TYPE "ST_StepRecord"
VERSION : 0.1
   STRUCT
      "StepNo" : Int;
      "StepName" : String[120];
      "AwaitingLabel" : String[120];
      "TimeClass" : DInt;
      "ExpectedTime" : Time;
      "Conds" : Array[1..8] of "ST_CondRecord";
   END_STRUCT;
END_TYPE
